Universal Robots URScript: T013_mistralai_Devstral-Small-2-24B-Instruct-2512_baseline_rep1.urscript

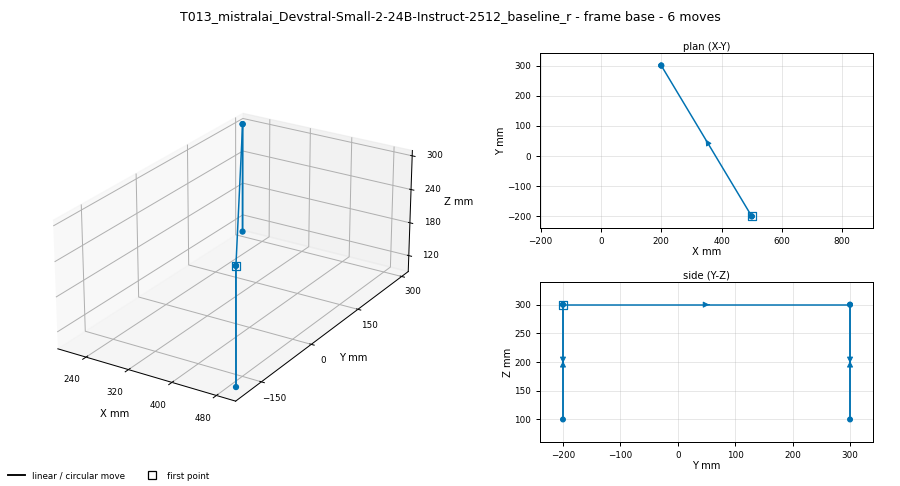
[picture p0: tool path of T013_mistralai_Devstral-Small-2-24B-Instruct-2512_baseline_rep1.urscript in frame base, 6 of 8 moves have a stored position in this frame; points joined in program order, loops and branches not executed]
def palletize_light_boxes():
    # Home position
    movej([0, -1.57, 0, -1.57, 0, 0], a=1.35, v=0.2, t=0, r=0)

    # Above staging area
    movel(p[0.5, -0.2, 0.3, 0, 3.14, 0], a=1.35, v=0.22, t=0, r=0)

    # Descend to pick
    movel(p[0.5, -0.2, 0.1, 0, 3.14, 0], a=1.35, v=0.1, t=0, r=0)

    # Lift
    movel(p[0.5, -0.2, 0.3, 0, 3.14, 0], a=1.35, v=0.18, t=0, r=0)

    # Transit to pallet
    movel(p[0.2, 0.3, 0.3, 0, 3.14, 0], a=1.35, v=0.23, t=0, r=0)

    # Descend to place
    movel(p[0.2, 0.3, 0.1, 0, 3.14, 0], a=1.35, v=0.1, t=0, r=0)

    # Lift after placing
    movel(p[0.2, 0.3, 0.3, 0, 3.14, 0], a=1.35, v=0.18, t=0, r=0)

    # Return to home
    movej([0, -1.57, 0, -1.57, 0, 0], a=1.35, v=0.2, t=0, r=0)

    # Safety zone confinement
    set_safety_zone_confinement(True)
